// TIA Portal V20 export
TYPE "DATA_RECEPT"
   STRUCT
      NUMBER_PROG { S7_SetPoint := 'True'} : Int;
      PROG_NAME { S7_SetPoint := 'True'} : String[38];
      OS_Z { S7_SetPoint := 'True'} : DInt;
      SELECTED : Bool;
   END_STRUCT;
END_TYPE
